(* IEC 61131-3 sources: plc-workbench/reports/tia_final_20261104/pairs/alias, 1 file *)

(* ---- baseline.st ---- *)
FUNCTION_BLOCK Demo
VAR_INPUT x : DINT; END_VAR
VAR_OUTPUT y : DINT; END_VAR
VAR_IN_OUT a : ARRAY[*] OF DINT; b : DINT; END_VAR
VAR copyDone : BOOL; idx : DINT; END_VAR
a[LOWER_BOUND(a, 1)] := x; y := b;
END_FUNCTION_BLOCK
